TYPE ST_VC_MoveToPositionResult :
STRUCT
    Accepted : BOOL;
END_STRUCT
END_TYPE

(* stored: Version 1.1.0.1, ProductVersion 3.1.4026.21
   DUT ST_VC_MoveToPositionResult: Id {5d2faee6-b6e3-4f14-ae49-713524515a1d} *)
